FUNCTION_BLOCK MicroswitchCheck
VAR_INPUT
END_VAR
VAR_OUTPUT
END_VAR
VAR
	SwTheta1: BOOL;
	SwTheta2: BOOL;
	SwR1: BOOL;
	SwR2: BOOL;
	SwBeta1: BOOL;
	SwBeta2: BOOL;
END_VAR

SwTheta1 	 := (GVL_MicroSwitch.dwMicroSwitchDriverA AND 16#00020000) <> 0;  (* bit 0 *)
SwTheta2     := (GVL_MicroSwitch.dwMicroSwitchDriverA AND 16#00010000) <> 0;  (* bit 1 *)
SwR1    	 := (GVL_MicroSwitch.dwMicroSwitchDriverB AND 16#00080000) <> 0;  (* bit 0 *)
SwR2  		 := (GVL_MicroSwitch.dwMicroSwitchDriverB AND 16#00040000) <> 0;  (* bit 1 *)
SwBeta1      := (GVL_MicroSwitch.dwMicroSwitchDriverB AND 16#00020000) <> 0;  (* bit 2 *)
SwBeta2      := (GVL_MicroSwitch.dwMicroSwitchDriverB AND 16#00010000) <> 0;  (* bit 3 *)

IF SwTheta1 THEN
GVL_HMI.CheckMicroswitchWristLeft := TRUE;
	
END_IF

IF SwTheta2 THEN
GVL_HMI.CheckMicroswitchWristRight := TRUE;
	
END_IF

IF SwR1 THEN
GVL_HMI.CheckMicroswitchLinearMax := TRUE;
	
END_IF

IF SwR2 THEN
GVL_HMI.CheckMicroswitchLinearMin := TRUE;
	
END_IF

IF SwBeta1 THEN
GVL_HMI.CheckMicroswitchRotationRight := TRUE;
	
END_IF

IF SwBeta2 THEN
GVL_HMI.CheckMicroswitchRotationLeft := TRUE;
	
END_IF

IF GVL_HMI.CheckMicroswitchWristLeft AND GVL_HMI.CheckMicroswitchWristRight AND GVL_HMI.CheckMicroswitchLinearMax AND GVL_HMI.CheckMicroswitchLinearMin AND GVL_HMI.CheckMicroswitchRotationRight AND GVL_HMI.CheckMicroswitchRotationLeft THEN
GVL_HMI.ContinueToHoming := TRUE;

END_IF

END_FUNCTION_BLOCK

(* stored: Version 1.1.0.1, ProductVersion 3.1.4024.15
   POU MicroswitchCheck: Id {1c0e4854-5048-4d36-942b-b7de663fad62}, SpecialFunc None *)
